(* CODESYS project GeneralControls.xml

Project tree, tasks and I/O mapping:
  visualisation GeneralControls
*)

// /GeneralControls
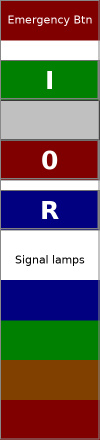
VISUALIZATION GeneralControls  // 100x440
    Rectangle (0,100 100x40), colour toggle: GVL_Project.fbProject._fbGeneralController._xSignalLightStartBtn
    Rectangle (0,320 100x40), colour toggle: GVL_Project.fbProject._fbGeneralController._xSignalLightGreen
    Rectangle (0,360 100x40), colour toggle: GVL_Project.fbProject._fbGeneralController._xSignalLightOrange
    Rectangle (0,400 100x40), colour toggle: GVL_Project.fbProject._fbGeneralController._xSignalLightRed
    Button (0,60 100x40), "I"
        tap GVL_Project.fbProject._fbGeneralController._btnStart.xbtn
    Button (0,140 100x40), "0"
        tap GVL_Project.fbProject._fbGeneralController._btnStop.xbtn
    Label (0,240 100x40), "Signal lamps"
    Rectangle (0,0 100x40), "Emergency Btn", colour toggle: GVL_Project.fbProject._fbGeneralController._xEmergencyBtnState
    Rectangle (0,280 100x40), colour toggle: GVL_Project.fbProject._fbGeneralController._xSignalLightResetBtn
    Button (0,190 100x40), "R"
        tap GVL_Project.fbProject._fbGeneralController._btnReset.xbtn
END_VISUALIZATION
